Fanuc KAREL source: kt00158.KL

-- PROVISIONAL review KL for V940-1; original PC SHA256 8039314fae67524e4e0117a7e6e8cbc8ce4b750fa4cb430957773e983310fedf
-- Incomplete behavior may be omitted. Consult companion uncertainty JSON. Do not deploy.
PROGRAM KT00158
%NOLOCKGROUP
VAR
  OUT : REAL
-- UNRESOLVED_DECL H1 type=002017
-- UNRESOLVED_DECL Y2 type=002018
BEGIN
  -- V9_ZERO_TABLE_METADATA_HINT layout=0001; no indexed target words; source/name/runtime held
  -- UNRESOLVED_PC offsets 5-19; opcodes 2E,22,9D,33,B4
  -- UNRESOLVED_PC offsets 24-38; opcodes 2E,22,9D,33,B2
  -- UNRESOLVED_PC offsets 43-69; opcodes 22,9D,33,B3,22,9D,33,B1,55,64,23
  -- UNRESOLVED_PC offsets 74-78; opcodes 7F
END KT00158
